(* IEC 61131-3 sources: rusty/compiler/plc_cfc/fixtures/blocks/valid/program_cycle, 1 file *)

(* ---- callees.st ---- *)
PROGRAM ping
VAR_INPUT
    in : DINT;
END_VAR
VAR_OUTPUT
    out : DINT;
END_VAR
    out := in + 1;
END_PROGRAM

PROGRAM pong
VAR_INPUT
    in : DINT;
END_VAR
VAR_OUTPUT
    out : DINT;
END_VAR
    out := in + 1;
END_PROGRAM
